(* IEC 61131-3 sources: ISA-88-Bioreactor-Automation-Template-DE-IE/ISA-88-Bioreactor-Automation-Template-DE-IE.fbsdev/PumpController.iecapp^/FunctionBlock, 4 files *)

(* ---- PumpAlarm_FB_ST.fb.st ---- *)
FUNCTION_BLOCK PumpAlarm_FB_ST
VAR_INPUT
    Pump_Discharge : BOOL;   // pump running
    Tn_Level_Low   : BOOL;   // tank empty sensor
    PT             : TIME := T#5s; // timeout duration
END_VAR

VAR_OUTPUT
    Pump_Alarm : BOOL := FALSE;
END_VAR

VAR
    TON_Alarm : TON; // IEC timer instance
END_VAR

// Alarm logic
IF Pump_Discharge AND NOT Tn_Level_Low THEN
    TON_Alarm(IN := TRUE, PT := PT);
ELSE
    TON_Alarm(IN := FALSE, PT := PT);
    Pump_Alarm := FALSE;
END_IF;

IF TON_Alarm.Q THEN
    Pump_Alarm := TRUE;
END_IF;

(* ---- PumpCycling_FB_ST.fb.st ---- *)
FUNCTION_BLOCK PumpController_FB_ST
VAR_INPUT
    Cycle_Active     : BOOL;   // cycle running
    Stage_Ready      : BOOL;   // stage condition met
    Tn_Level_Low     : BOOL;   // tank empty sensor
END_VAR

VAR_OUTPUT
    Pump_Discharge   : BOOL := FALSE;
    Discharge_Complete : BOOL := FALSE;
END_VAR

// Pump control logic
IF Cycle_Active AND Stage_Ready THEN
    Pump_Discharge := NOT Tn_Level_Low;
    IF Tn_Level_Low THEN
        Discharge_Complete := TRUE;
        Pump_Discharge := FALSE;
    END_IF;
ELSE
    Pump_Discharge := FALSE;
    Discharge_Complete := FALSE;
END_IF;

(* ---- PumpInterlock_FB_ST.fb.st ---- *)
FUNCTION_BLOCK PumpInterlock_FB_ST
VAR_INPUT
    Heater : BOOL; // heater ON/OFF
END_VAR

VAR_OUTPUT
    Pump_Enable : BOOL := FALSE;
END_VAR

// Interlock logic
Pump_Enable := NOT Heater;

(* ---- PumpTimer_FB_ST.fb.st ---- *)
FUNCTION_BLOCK PumpTimer_FB_ST
VAR_INPUT
    Cycle_Active : BOOL;   // overall cycle running
    Stage_Ready  : BOOL;   // discharge stage condition met
    PT           : TIME := T#10s; // preset time (adjust as needed)
END_VAR

VAR_OUTPUT
    PumpTimer_Done : BOOL := FALSE;
END_VAR

VAR
    TON_Pump : TON; // IEC timer instance
END_VAR

// Timer logic
TON_Pump(IN := (Cycle_Active AND Stage_Ready), PT := PT);

PumpTimer_Done := TON_Pump.Q;
